(*
    This function runs all test suites that have been initialized.
    The test suites are run in sequence (one after the other).
*)
FUNCTION RUN_IN_SEQUENCE

GVL_TcUnit.TcUnitRunner.RunTestSuiteTestsInSequence(TimeBetweenTestSuitesExecution := GVL_Param_TcUnit.TimeBetweenTestSuitesExecution);

END_FUNCTION

(* stored: Version 1.1.0.1
   POU RUN_IN_SEQUENCE: Id {a1bb30cd-f92f-4bab-aa26-6bd18db0fbc1}, SpecialFunc None *)
